// TIA Portal V20 export
// export: Created 2026-10-19T18:06:46.3339109Z, ExportSetting WithDefaults, DisplayName Totally Integrated Automation Portal, DisplayVersion V20 Update 6, DisplayName TIA Portal Openness, DisplayVersion V20 Update 6, DisplayName TIA Portal Version Control Interface, DisplayVersion V20 Update 6, DisplayName SINAMICS Startdrive Advanced, DisplayVersion V20 SP1, DisplayName SINAMICS Startdrive G130, G150, S120, S150, SINAMICS MV, G220, S200, S210, DisplayVersion V20 SP1, DisplayName SINAMICS Startdrive G110M, G120, G120C, G120D, G120P, G115D, DisplayVersion V20 SP1, DisplayName STEP 7 Professional, DisplayVersion V20 Update 6, DisplayName STEP 7 Safety, DisplayVersion V20 Update 2, DisplayName WinCC Basic/Comfort/Advanced, DisplayVersion V20 Update 6, DisplayName WinCC Unified, DisplayVersion V20 Update 6
DATA_BLOCK "SAI_IND_AlibiRead_DB"   // DB107
VERSION : 0.1
// stored: AutoNumber true, DBAccessibleFromOPCUA true, DBAccessibleFromWebserver true, InstanceOfName SAI_IND360Base_AlibiRead, InstanceOfType FB
"SAI_IND360Base_AlibiRead"
   // VAR_INPUT
   //    ID : HW_IO;
   // END_VAR
   // VAR_OUTPUT
   //    Done : Bool;
   //    Error : Bool;
   //    GrossWeight : Real;
   //    TareWeight : Real;
   //    NetWeight : Real;
   //    TareMode : SInt;
   //    Unit : SInt;
   // END_VAR
   // VAR_IN_OUT
   //    ePrint : Bool;
   //    RecordNumber : DInt;
   //    Get_TransactionNum : Bool;
   //    Set_TransactionNum : Bool;
   //    Get_Alibi : Bool;
   //    Alibi_Array : Array[0..44] of Byte;
   // END_VAR
   // VAR
   //    RDREC01 { S7_SetPoint := 'True'} : RDREC;
   //    RDREC02 { S7_SetPoint := 'True'} : RDREC;
   //    WRREC01 { S7_SetPoint := 'True'} : WRREC;
   //    WRREC02 { S7_SetPoint := 'True'} : WRREC;
   //    UINT : SInt;
   // END_VAR
BEGIN
END_DATA_BLOCK
